TYPE ET_STOEBER_AxisSetLimitsTc2 :
(
	ET_STOEBER_AxisSetLimits_eWaitExecute := 0,
	ET_STOEBER_AxisSetLimits_eSetLimitPos,
	ET_STOEBER_AxisSetLimits_eSetLimitNeg,
	ET_STOEBER_AxisSetLimits_eSetJogVelo,
	ET_STOEBER_AxisSetLimits_eSetJogAcc,
	ET_STOEBER_AxisSetLimits_eSetJogDec,
	ET_STOEBER_AxisSetLimits_eSetJogJerk,
	ET_STOEBER_AxisSetLimits_eDone := 197,
	ET_STOEBER_AxisSetLimits_eError := 198,
	ET_STOEBER_AxisSetLimits_eNoExecute := 199
);
END_TYPE

(* stored: Version 1.1.0.1, ProductVersion 3.1.4024.15
   DUT ET_STOEBER_AxisSetLimitsTc2: Id {1c90c5a2-724f-4550-bd5c-b763c21af256} *)
